(* IEC 61131-3 sources: kns-port-domestic/targets/astra/lib/src/DUTs/DigitalInput, 5 files *)

(* ---- E_DiAlarm.dut.st ---- *)
// Назначение: индексы слотов тревог дискретного входа. Нестрогое перечисление: им
//             индексируются массивы.
// Автор:      kr0nsch
// Версия:     0.1.0
// Документ:   docs/fb/FB_DigitalInput.md
{attribute 'qualified_only'}
TYPE E_DiAlarm :
(
    State   := 0,   // тревога по состоянию сигнала (включает генератор, если сигнал тревожный)
    Failure := 1    // отказ канала
) UINT;
END_TYPE

(* ---- E_DiFailValue.dut.st ---- *)
// Назначение: значение дискретного входа при отказе канала.
// Автор:      kr0nsch
// Версия:     0.1.0
// Документ:   docs/fb/FB_DigitalInput.md
{attribute 'qualified_only'}
{attribute 'strict'}
TYPE E_DiFailValue :
(
    HoldLast   := 0,   // удерживать последнее значение
    ForceFalse := 1,
    ForceTrue  := 2    // для защитных сигналов: отказ канала = сработал
) INT;
END_TYPE

(* ---- ST_DigitalInputCfg.dut.st ---- *)
// Назначение: параметры дискретного входа (Persistent Variables приложения,
//             VAR_IN_OUT CONSTANT stCfg). Значения по умолчанию проходят CheckConfig.
//             Тип лежит в Persistent Variables приложения и заморожен в пределах 1.x (A-13).
// Автор:      kr0nsch
// Версия:     0.1.0
// Документ:   docs/fb/FB_DigitalInput.md
{attribute 'qualified_only'}
TYPE ST_DigitalInputCfg :
STRUCT
    xInvert        : BOOL := FALSE;    // инверсия до задержек (НЗ-контакт)
    tOnDelay       : TIME := T#0S;     // задержка включения
    tOffDelay      : TIME := T#0S;     // задержка отключения
    eFailValue     : E_DiFailValue := E_DiFailValue.HoldLast;
    xAlarmOnTrue   : BOOL := TRUE;     // тревога State при xValue = TRUE (FALSE — при xValue = FALSE)
    tSubstMax      : TIME := T#8H;     // макс. длительность подмены; T#0S — без ограничения
    udiAlarmIdBase : UDINT := 0;       // номер первой тревоги устройства (dev_no * 10)
    astAlarm       : ARRAY[0..GVL_Const.DEV_ALARMS_MAX - 1] OF ST_AlarmCfg := [
        (ePriority := E_AlarmPriority.None),      // 0 State — включает генератор, если сигнал тревожный
        (ePriority := E_AlarmPriority.Medium),    // 1 Failure
        (ePriority := E_AlarmPriority.None), (ePriority := E_AlarmPriority.None),
        (ePriority := E_AlarmPriority.None), (ePriority := E_AlarmPriority.None),
        (ePriority := E_AlarmPriority.None), (ePriority := E_AlarmPriority.None)];
END_STRUCT
END_TYPE

(* ---- ST_DigitalInputCmd.dut.st ---- *)
// Назначение: команды HMI/SCADA дискретного входа (GVL_Hmi приложения, VAR_IN_OUT stCmd).
// Автор:      kr0nsch
// Версия:     0.1.0
// Документ:   docs/fb/FB_DigitalInput.md
{attribute 'qualified_only'}
TYPE ST_DigitalInputCmd :
STRUCT
    stCommon    : ST_DeviceCmd;   // xSetAuto — «Измерение», xSetManual — «Подмена»
    xSubstValue : BOOL;           // значение подмены; в Auto ФБ пишет сюда текущее xValue
END_STRUCT
END_TYPE

(* ---- ST_DigitalInputSts.dut.st ---- *)
// Назначение: состояние дискретного входа для HMI/SCADA. 30 байт, 15 регистров Modbus.
//             Значение и сырой сигнал — биты DI_STS_VALUE / DI_STS_RAW в stCommon.wStatus и выход
//             экземпляра xValue: полей BOOL в Sts нет.
// Автор:      kr0nsch
// Версия:     0.1.0
// Документ:   docs/fb/FB_DigitalInput.md
{attribute 'qualified_only'}
TYPE ST_DigitalInputSts :
STRUCT
    stCommon        : ST_DeviceSts;   // 0..27
    uiSubstRemain_s : UINT;           // 28: до автоматического снятия подмены, с; 0 — подмены нет
END_STRUCT
END_TYPE
